Fanuc KAREL source: KO00056.KL

PROGRAM KO00056
%NOLOCKGROUP
%ENVIRONMENT MIR
VAR
  P1: XYZWPR
  P2: XYZWPR
  F: BOOLEAN
  OUT: JOINTPOS
BEGIN
  F = TRUE
  OUT = MIRROR(P1, P2, F)
END KO00056
